Fanuc KAREL source: KA00034.KL

PROGRAM KA00034
%NOLOCKGROUP
VAR
  SRC: BOOLEAN
  DST: CONFIG
BEGIN
  SRC = TRUE
  DST = SRC
END KA00034
